(* IEC 61131-3 sources: plcassist-cli/packages/volt-lsp-iec/test-corpus/bakon-nano/Device/Plc Logic/Application/Library Manager/CmpSrv, 2 files *)

(* ---- COMPONENTID.gvl ---- *)
VAR_GLOBAL
	CMPID_CMPSRV : UDINT := 16#1C;
END_VAR

(* ---- EVENTIDS.gvl ---- *)
VAR_GLOBAL
	EVTPARAMID_CMPSRV : UDINT := 16#1;
	EVTVERSION_CMPSRV : UDINT := 16#2;
END_VAR
